(* Logix 5000 project; controller TFF vendor 1 type 14 code 107 rev 34.11; software revision 34.03; part 28 of 36 *)
(* tags used below, declared in another part *)
   Config : Configuration;   // Index Array used in configuration routines
   AlarmControl : AlarmControl;   // Alarm Control
   AnalogOutput : AnalogOutput[25];   // Analog Output Array
   AnalogPoint : AnalogInput[50];   // Analog Input Array
   CCPSystem : CCPSystem;   // CCP System Data
   ChartMark : ChartMark;   // Chart Mark
   Concentration : Concentration;
   CPU_Scanning : BOOL;   // System Scanning Flag
   Diafiltration : Diafiltration;
   DigitalOutput : BOOL[256];   // Digital Output Array these bits are sent to output cards.
   DigitalPoint : DigitalPoint[150];   // Digital Point Array
   DPAlarm : ALIAS FOR AlarmAnalog[40];   // Differential Pressure Alarm
   Drive : Drive[11];   // Drives Array
   ES001 : ALIAS FOR DigitalPoint[3];   // Emergency Stop
   Feed_Pump_P001_Type : INT;   // Feed Pump P001 Type Status
   FirstScanComplete : BOOL;   // First Scan Complete Flag
   FlowPath : FlowPath[64];   // Flow Path Array
   Membrane_Data : Membrane_Data;   // Membrane Data
   Mixer : Mixer;   // Mixer config. structure
   OperatingTime : OperatingTime;
   Operation : Operation[6,251];   // Operation Table
   Options : Options;   // Options List
   Phase0 : ALIAS FOR Phase[0];   // Phase 0
   Phase0_Totalizer_Feed : ALIAS FOR PhaseTotalizer[0];   // Phase 0 Total Feed
   Phase0_Totalizer_Filtrate : ALIAS FOR PhaseTotalizer[6];   // Phase 0 Total Filtrate
   Phase0_Totalizer_Retentate : ALIAS FOR PhaseTotalizer[12];   // Phase 0 Total Retentate
   PipeAnimation : PipeAnimation;   // HMI Pipe Animation Array
   PLCFault : FaultRecordType;   // PLC Major Fault Record
   PumpRunStatus : DINT;   // Pumps Run Status (1 = At least one pump running , 0 = no pump running)
   Rack_Murr_Node6_IND331_WI001 : IO_Station;   // Status of Node 6 IND331 WI001
   Rack_Murr_Node7_IND131_WI101 : IO_Station;   // Status of Node 7 IND131 WI101
   SIC001 : ALIAS FOR Drive[1];   // Feed Pump
   SIC002 : ALIAS FOR Drive[2];   // Transfer Pump
   SIC003 : ALIAS FOR Drive[3];   // Mixer
   SIC003DF : ALIAS FOR DigitalPoint[14];   // Mixer Defect
   SysControl : SysControl;   // General system status and command
   Tank : TankManagement;   // Tank Management
   ThisSystem : SystemType;
   TimerControl : TimerControl;   // Timer Control
   Timers : Timers[22];   // Timer Array
   TMPAlarm : ALIAS FOR AlarmAnalog[41];   // Trans-membrane Pressure Alarm
   Totalizer : Totalizers[20];   // Totalizers Array
   Transfer_Pump_P002_Type : INT;   // Transfer Pump P002 Type Status
   UserAlarm : UserAlarm;   // User Alarm (used in CCP Recipe)
   UserCr1 : ALIAS FOR DigitalPoint[65];   // User Critical Alarm 1
   UserCr2 : ALIAS FOR DigitalPoint[67];   // User Critical Alarm 2
   UserNCr1 : ALIAS FOR DigitalPoint[64];   // User Non Critical Alarm 1
   UserNCr2 : ALIAS FOR DigitalPoint[66];   // User Non Critical Alarm 2
   UserTime : ALIAS FOR Timers[18];   // User time
   UserTotalizerManagement : UserTotalizerManagement;   // User Totalizer management
   Valve : Valve[100];   // Valve Array
   XC102_3 : ALIAS FOR DigitalOutput[5];   // UV Auto Zero
   XS011 : ALIAS FOR DigitalPoint[11];   // Pump P001 Type
   XS012 : ALIAS FOR DigitalPoint[12];   // Pump P002 Type
   YA10 : ALIAS FOR DigitalPoint[59];   // PLC Program Major Fault
   YA41 : ALIAS FOR DigitalPoint[77];   // YA41 Operating Time Exceeded
(* Process, continued *)

ROUTINE InputProcessing   (* ladder *)
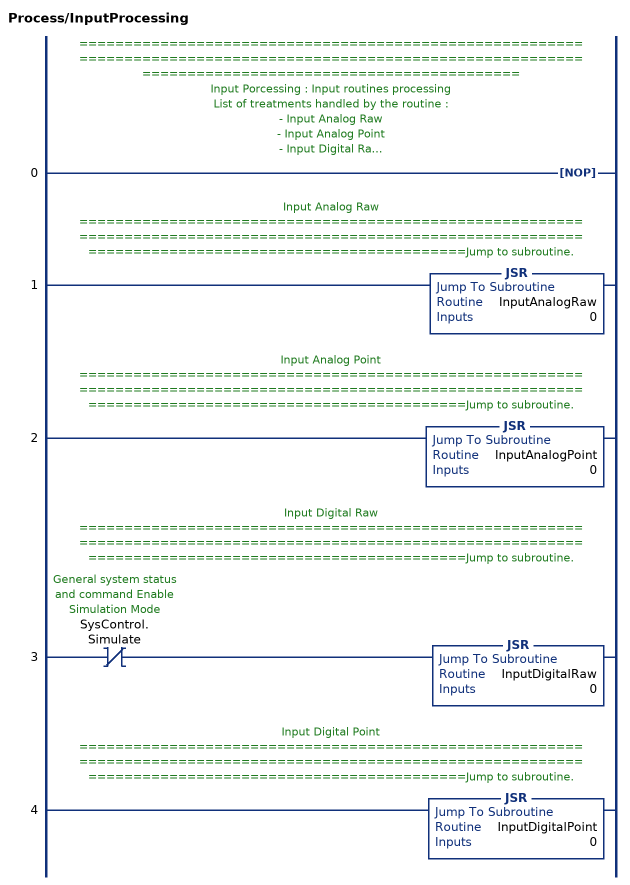
   // ==========================================================================================================================================================
   //                                                                                                                      Input Porcessing : Input routines processing
   //                                                     List of treatments handled by the routine :
   //                                                          - Input Analog Raw
   //                                                          - Input Analog Point
   //                                                          - Input Digital Raw
   //                                                          - Input Digital Point
   //                                                     -----------------------------------------------------------------------------------------------------------------------------------------------------
   //                                                     History
   //                                                          2019-AUG-13 - Actemium - B. Roch - Initial version for Candidate Release 3.00.00.00.a
   // ==========================================================================================================================================================
   0: NOP();
   // Input Analog Raw
   // ==========================================================================================================================================================Jump to subroutine.
   1: JSR(InputAnalogRaw,0);
   // Input Analog Point
   // ==========================================================================================================================================================Jump to subroutine.
   2: JSR(InputAnalogPoint,0);
   // Input Digital Raw
   // ==========================================================================================================================================================Jump to subroutine.
   3: XIO(SysControl.Simulate)JSR(InputDigitalRaw,0);
   // Input Digital Point
   // ==========================================================================================================================================================Jump to subroutine.
   4: JSR(InputDigitalPoint,0);
END_ROUTINE

ROUTINE MainRoutine   (* ladder *)
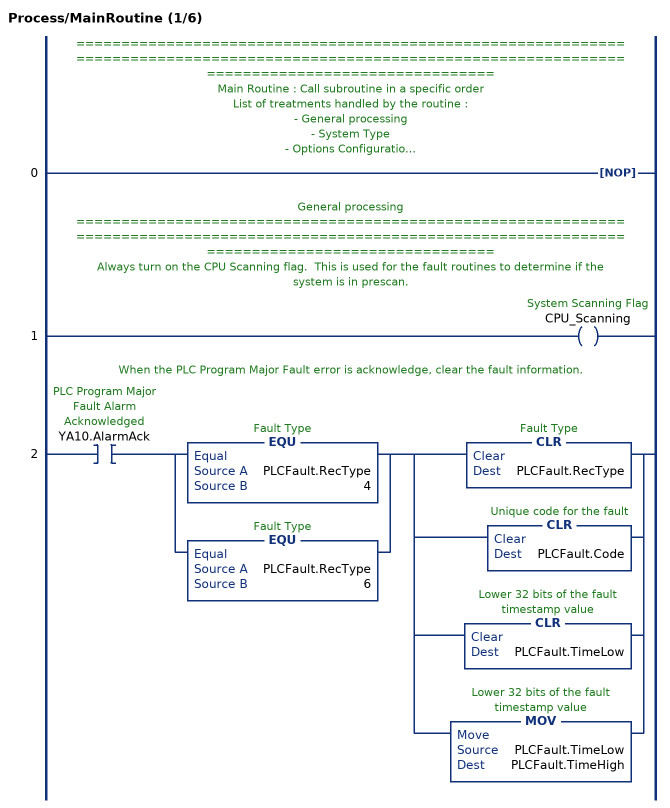
   // ==========================================================================================================================================================
   //                                                                                                            Main Routine : Call subroutine in a specific order
   //                                                     List of treatments handled by the routine :
   //                                                          - General processing
   //                                                          - System Type
   //                                                          - Options Configuration
   //                                                          - AnalogOutput Configuration
   //                                                          - AnalogPoint Configuration
   //                                                          - DigitalPoint Configuration (real input)
   //                                                          - DigitalPoint Configuration (soft input)
   //                                                          - Valve Configuration
   //                                                          - Drive Configuration
   //                                                          - Control Loop Configuration
   //                                                          - Totalizers Configuration
   //                                                          - Flowpath Configuration
   //                                                          - Reset Configuration
   //                                                          - Station Status
   //                                                          - Derived Data
   //                                                          - Analog and Digital Input Processing
   //                                                          - Pump Control
   //                                                          - Loop Control
   //                                                          - Valve Control
   //                                                          - Pipe Animation
   //                                                          - Alarm
   //                                                          - Concentration & Diafiltration
   //                                                          - TankManagement
   //                                                          - Miscellaneous Functions
   //                                                          - Analog and Digital Output Processing
   //                                                     -----------------------------------------------------------------------------------------------------------------------------------------------------
   //                                                     History
   //                                                          2019-AUG-13 - Actemium - B. Roch - Initial version for Candidate Release 3.00.00.00.a
   //                                                          2020-SEP-14 - Merck - Q. Spindler - Modifications for Candidate Release 3.00.00.01.a
   //                                                                  - Add TimerControl.TickMainTask for 1 sec tick in Main task
   // ==========================================================================================================================================================
   0: NOP();
   // General processing
   // ==========================================================================================================================================================
   // Always turn on the CPU Scanning flag.  This is used for the fault routines to determine if the system is in prescan.
   1: OTE(CPU_Scanning);
   // When the PLC Program Major Fault error is acknowledge, clear the fault information.
   2: XIC(YA10.AlarmAck)[EQU(PLCFault.RecType,4) ,EQU(PLCFault.RecType,6) ][CLR(PLCFault.RecType) ,CLR(PLCFault.Code) ,CLR(PLCFault.TimeLow) ,MOV(PLCFault.TimeLow,PLCFault.TimeHigh) ];
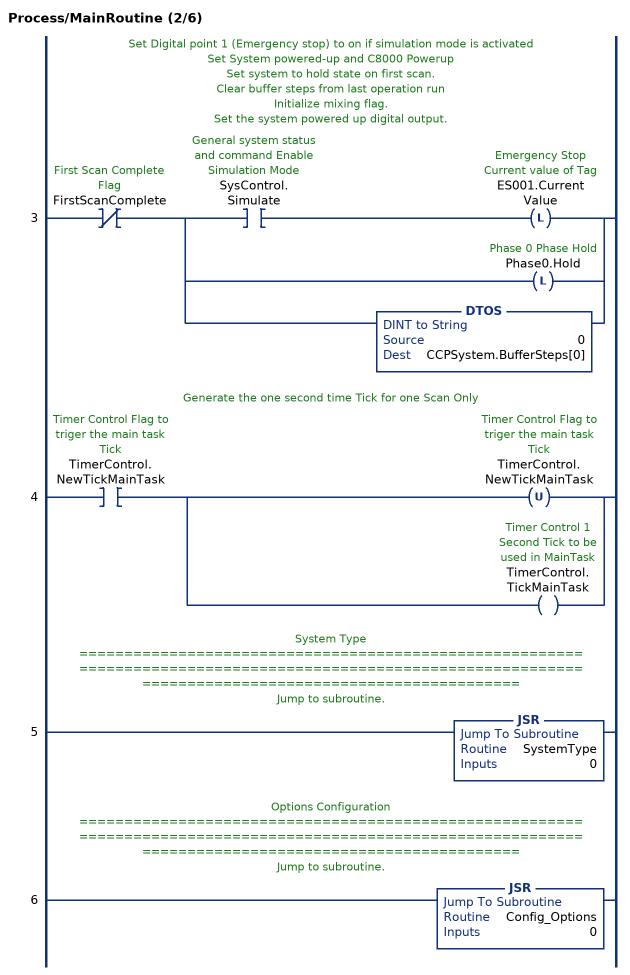
   // Set Digital point 1 (Emergency stop) to on if simulation mode is activated
   // Set System powered-up and C8000 Powerup
   // Set system to hold state on first scan.
   // Clear buffer steps from last operation run
   // Initialize mixing flag.
   // Set the system powered up digital output.
   3: XIO(FirstScanComplete)[XIC(SysControl.Simulate) OTL(ES001.CurrentValue) ,OTL(Phase0.Hold) ,DTOS(0,CCPSystem.BufferSteps[0]) ];
   // Generate the one second time Tick for one Scan Only
   4: XIC(TimerControl.NewTickMainTask)[OTU(TimerControl.NewTickMainTask) ,OTE(TimerControl.TickMainTask) ];
   // System Type
   // ==========================================================================================================================================================
   // Jump to subroutine.
   5: JSR(SystemType,0);
   // Options Configuration
   // ==========================================================================================================================================================
   // Jump to subroutine.
   6: JSR(Config_Options,0);
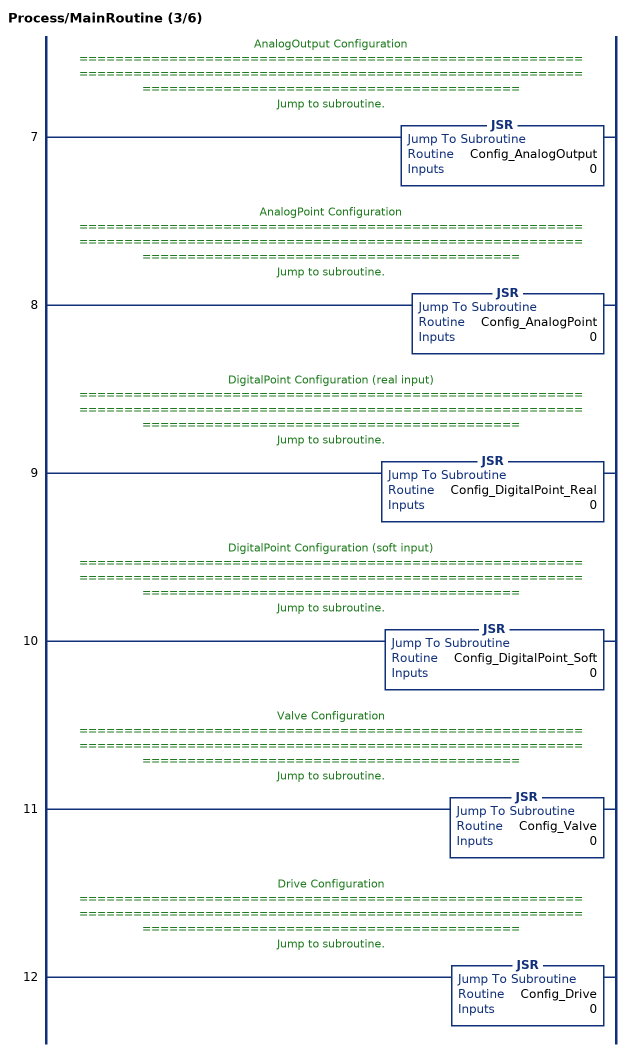
   // AnalogOutput Configuration
   // ==========================================================================================================================================================
   // Jump to subroutine.
   7: JSR(Config_AnalogOutput,0);
   // AnalogPoint Configuration
   // ==========================================================================================================================================================
   // Jump to subroutine.
   8: JSR(Config_AnalogPoint,0);
   // DigitalPoint Configuration (real input)
   // ==========================================================================================================================================================
   // Jump to subroutine.
   9: JSR(Config_DigitalPoint_Real,0);
   // DigitalPoint Configuration (soft input)
   // ==========================================================================================================================================================
   // Jump to subroutine.
   10: JSR(Config_DigitalPoint_Soft,0);
   // Valve Configuration
   // ==========================================================================================================================================================
   // Jump to subroutine.
   11: JSR(Config_Valve,0);
   // Drive Configuration
   // ==========================================================================================================================================================
   // Jump to subroutine.
   12: JSR(Config_Drive,0);
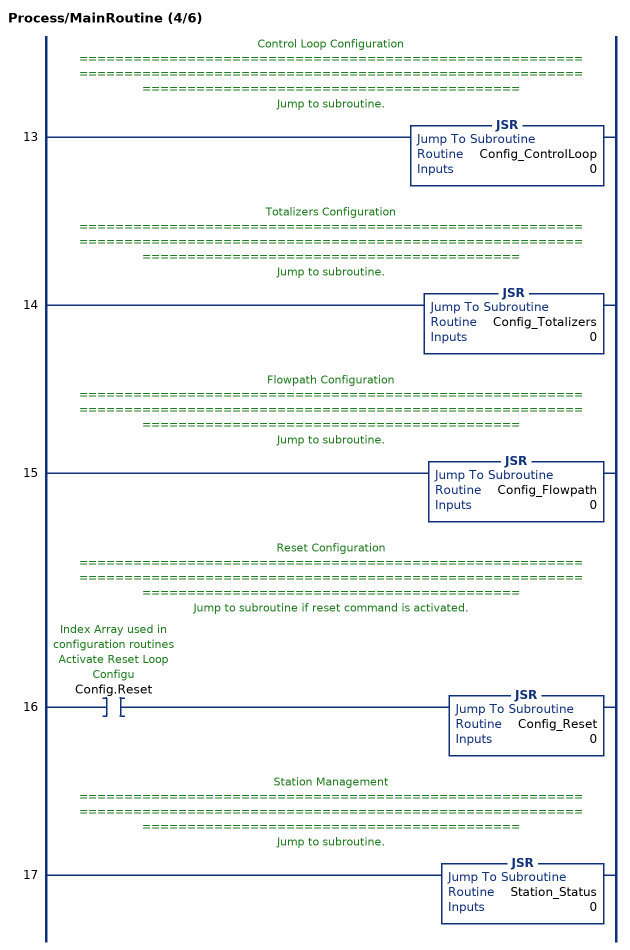
   // Control Loop Configuration
   // ==========================================================================================================================================================
   // Jump to subroutine.
   13: JSR(Config_ControlLoop,0);
   // Totalizers Configuration
   // ==========================================================================================================================================================
   // Jump to subroutine.
   14: JSR(Config_Totalizers,0);
   // Flowpath Configuration
   // ==========================================================================================================================================================
   // Jump to subroutine.
   15: JSR(Config_Flowpath,0);
   // Reset Configuration
   // ==========================================================================================================================================================
   // Jump to subroutine if reset command is activated.
   16: XIC(Config.Reset)JSR(Config_Reset,0);
   // Station Management
   // ==========================================================================================================================================================
   // Jump to subroutine.
   17: JSR(Station_Status,0);
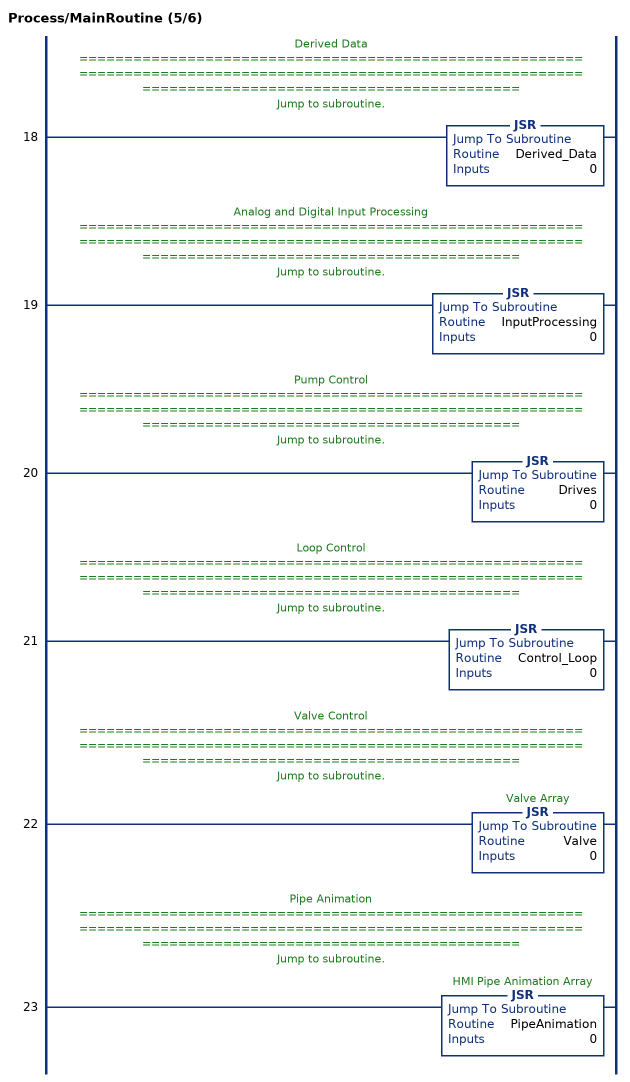
   // Derived Data
   // ==========================================================================================================================================================
   // Jump to subroutine.
   18: JSR(Derived_Data,0);
   // Analog and Digital Input Processing
   // ==========================================================================================================================================================
   // Jump to subroutine.
   19: JSR(InputProcessing,0);
   // Pump Control
   // ==========================================================================================================================================================
   // Jump to subroutine.
   20: JSR(Drives,0);
   // Loop Control
   // ==========================================================================================================================================================
   // Jump to subroutine.
   21: JSR(Control_Loop,0);
   // Valve Control
   // ==========================================================================================================================================================
   // Jump to subroutine.
   22: JSR(Valve,0);
   // Pipe Animation
   // ==========================================================================================================================================================
   // Jump to subroutine.
   23: JSR(PipeAnimation,0);
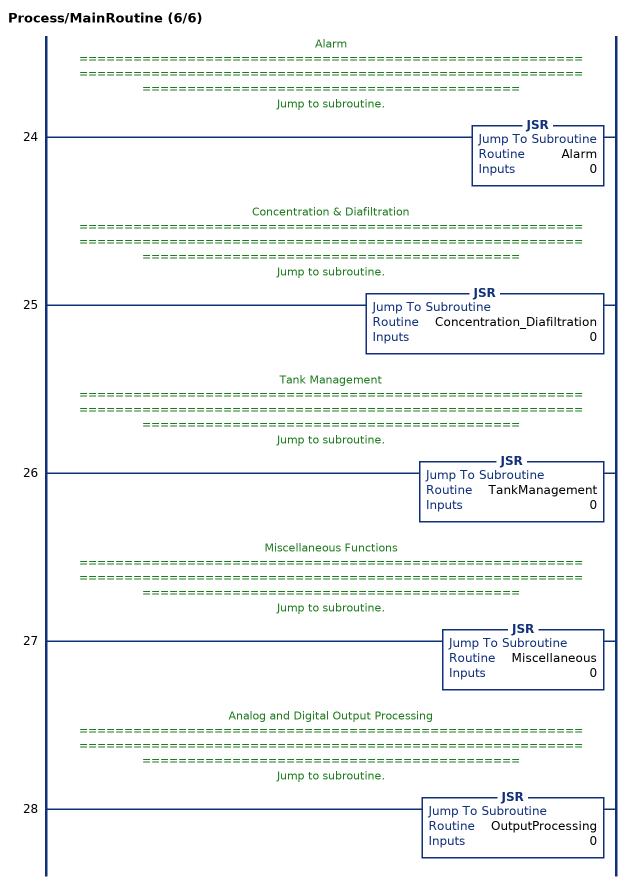
   // Alarm
   // ==========================================================================================================================================================
   // Jump to subroutine.
   24: JSR(Alarm,0);
   // Concentration & Diafiltration
   // ==========================================================================================================================================================
   // Jump to subroutine.
   25: JSR(Concentration_Diafiltration,0);
   // Tank Management
   // ==========================================================================================================================================================
   // Jump to subroutine.
   26: JSR(TankManagement,0);
   // Miscellaneous Functions
   // ==========================================================================================================================================================
   // Jump to subroutine.
   27: JSR(Miscellaneous,0);
   // Analog and Digital Output Processing
   // ==========================================================================================================================================================
   // Jump to subroutine.
   28: JSR(OutputProcessing,0);
END_ROUTINE

ROUTINE Miscellaneous   (* ladder *)
// Miscellaneous Routine
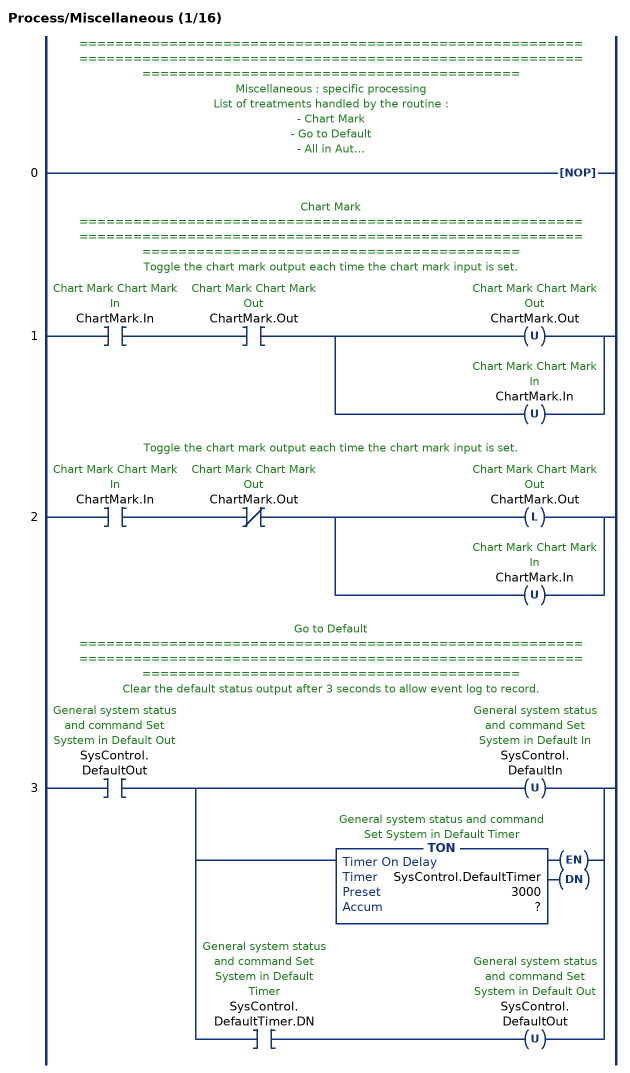
   // ==========================================================================================================================================================
   //                                                                                                                                 Miscellaneous : specific processing
   //                                                     List of treatments handled by the routine :
   //                                                          - Chart Mark
   //                                                          - Go to Default
   //                                                          - All in Auto
   //                                                          - Input Digital Point
   //                                                          - Enable All Alarms
   //                                                          - Disable All Alarms
   //                                                          - Enable all Analog signal alarms
   //                                                          - Disable all Analog signal alarms
   //                                                          - User totalizer management
   //                                                          - Pump Status calculation
   //                                                          - User Alarm (used in recipe only)
   //                                                          - Default Status
   //                                                          - Save \ Restore parameters conditions
   //                                                          - Mixer Reset Alarm Command
   //                                                          - IND331 and IND131 Configurations
   //                                                          - UV Baseline Zero Command Logic
   //                                                          - Pump Type Status
   //                                                     -----------------------------------------------------------------------------------------------------------------------------------------------------
   //                                                     History
   //                                                          2019-AUG-13 - Actemium - B. Roch - Initial version for Candidate Release 3.00.00.00.a
   //                                                          2019-OCT-25 - Actemium - B. Roch - Modification for Candidate Release 3.00.00.00.d
   //                                                         - Change Mixer Reset alarm condition SIC003DF.CurrentValue instead of SIC003DF.Alarm
   //                                                      2020-SEP-29 - Merck - Q. Spindler - Modifications for Candidate Release 3.00.00.01.a
   // 							- Add Retentate totalizer for UserTotalizer
   //                                                             2021-APR-30 - DAVIDSON- Ch. ARBOGAST - Modifications for Candidate Release 3.01.00.00.a
   //             -  Add Conditions to YA41 Operating Time Exceeded
   // ==========================================================================================================================================================
   0: NOP();
   // Chart Mark
   // ==========================================================================================================================================================
   // Toggle the chart mark output each time the chart mark input is set.
   1: XIC(ChartMark.In)XIC(ChartMark.Out)[OTU(ChartMark.Out) ,OTU(ChartMark.In) ];
   // Toggle the chart mark output each time the chart mark input is set.
   2: XIC(ChartMark.In)XIO(ChartMark.Out)[OTL(ChartMark.Out) ,OTU(ChartMark.In) ];
   // Go to Default
   // ==========================================================================================================================================================
   // Clear the default status output after 3 seconds to allow event log to record.
   3: XIC(SysControl.DefaultOut)[OTU(SysControl.DefaultIn) ,TON(SysControl.DefaultTimer,?,?) ,XIC(SysControl.DefaultTimer.DN) OTU(SysControl.DefaultOut) ];
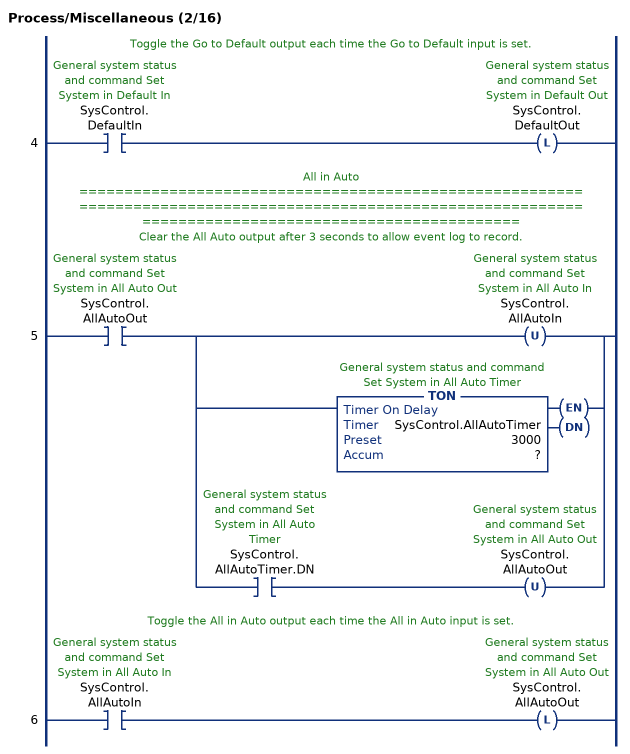
   // Toggle the Go to Default output each time the Go to Default input is set.
   4: XIC(SysControl.DefaultIn)OTL(SysControl.DefaultOut);
   // All in Auto
   // ==========================================================================================================================================================
   // Clear the All Auto output after 3 seconds to allow event log to record.
   5: XIC(SysControl.AllAutoOut)[OTU(SysControl.AllAutoIn) ,TON(SysControl.AllAutoTimer,?,?) ,XIC(SysControl.AllAutoTimer.DN) OTU(SysControl.AllAutoOut) ];
   // Toggle the All in Auto output each time the All in Auto input is set.
   6: XIC(SysControl.AllAutoIn)OTL(SysControl.AllAutoOut);
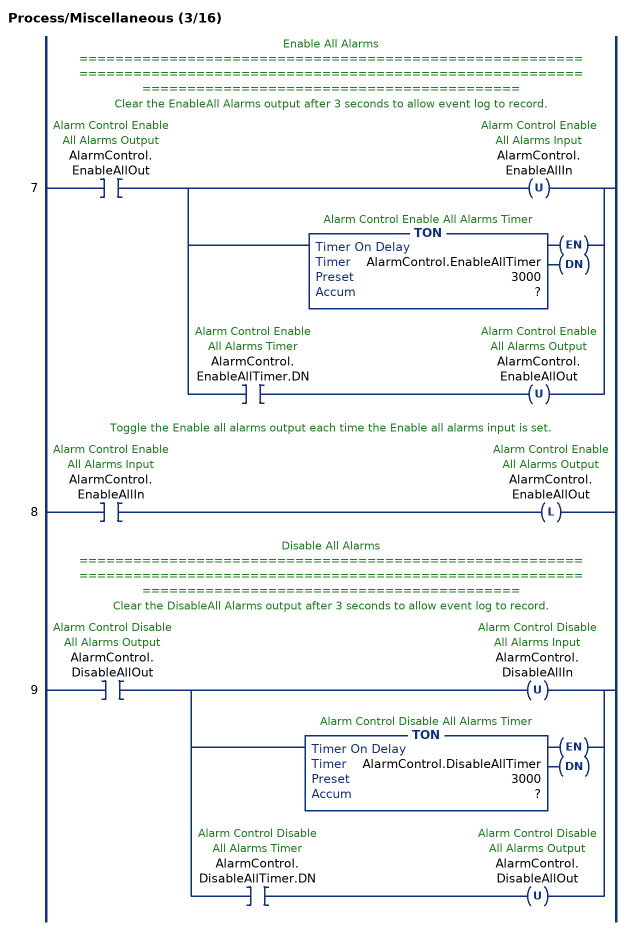
   // Enable All Alarms
   // ==========================================================================================================================================================
   // Clear the EnableAll Alarms output after 3 seconds to allow event log to record.
   7: XIC(AlarmControl.EnableAllOut)[OTU(AlarmControl.EnableAllIn) ,TON(AlarmControl.EnableAllTimer,?,?) ,XIC(AlarmControl.EnableAllTimer.DN) OTU(AlarmControl.EnableAllOut) ];
   // Toggle the Enable all alarms output each time the Enable all alarms input is set.
   8: XIC(AlarmControl.EnableAllIn)OTL(AlarmControl.EnableAllOut);
   // Disable All Alarms
   // ==========================================================================================================================================================
   // Clear the DisableAll Alarms output after 3 seconds to allow event log to record.
   9: XIC(AlarmControl.DisableAllOut)[OTU(AlarmControl.DisableAllIn) ,TON(AlarmControl.DisableAllTimer,?,?) ,XIC(AlarmControl.DisableAllTimer.DN) OTU(AlarmControl.DisableAllOut) ];
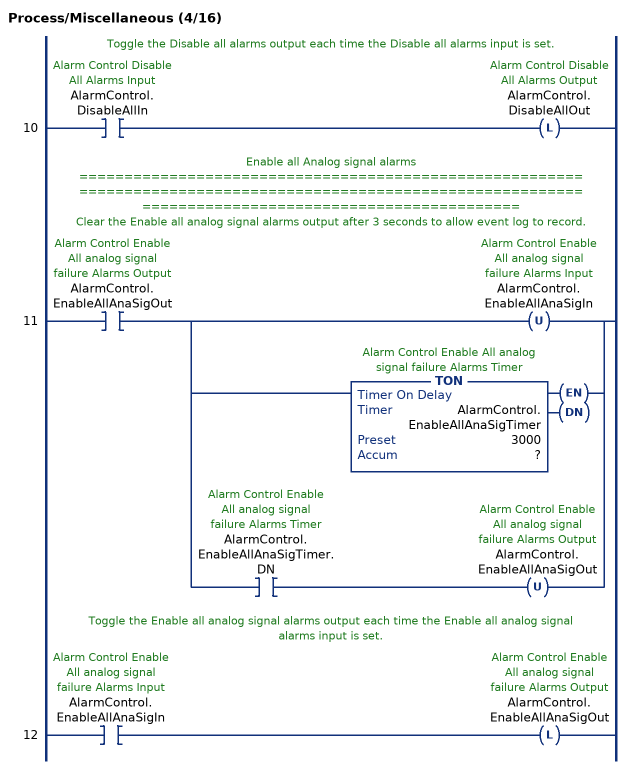
   // Toggle the Disable all alarms output each time the Disable all alarms input is set.
   10: XIC(AlarmControl.DisableAllIn)OTL(AlarmControl.DisableAllOut);
   // Enable all Analog signal alarms
   // ==========================================================================================================================================================
   // Clear the Enable all analog signal alarms output after 3 seconds to allow event log to record.
   11: XIC(AlarmControl.EnableAllAnaSigOut)[OTU(AlarmControl.EnableAllAnaSigIn) ,TON(AlarmControl.EnableAllAnaSigTimer,?,?) ,XIC(AlarmControl.EnableAllAnaSigTimer.DN) OTU(AlarmControl.EnableAllAnaSigOut) ];
   // Toggle the Enable all analog signal alarms output each time the Enable all analog signal alarms input is set.
   12: XIC(AlarmControl.EnableAllAnaSigIn)OTL(AlarmControl.EnableAllAnaSigOut);
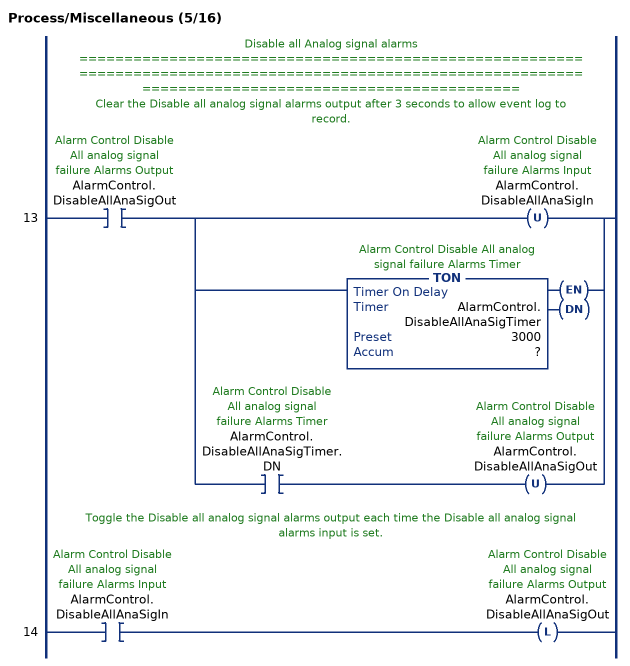
   // Disable all Analog signal alarms
   // ==========================================================================================================================================================
   // Clear the Disable all analog signal alarms output after 3 seconds to allow event log to record.
   13: XIC(AlarmControl.DisableAllAnaSigOut)[OTU(AlarmControl.DisableAllAnaSigIn) ,TON(AlarmControl.DisableAllAnaSigTimer,?,?) ,XIC(AlarmControl.DisableAllAnaSigTimer.DN) OTU(AlarmControl.DisableAllAnaSigOut) ];
   // Toggle the Disable all analog signal alarms output each time the Disable all analog signal alarms input is set.
   14: XIC(AlarmControl.DisableAllAnaSigIn)OTL(AlarmControl.DisableAllAnaSigOut);
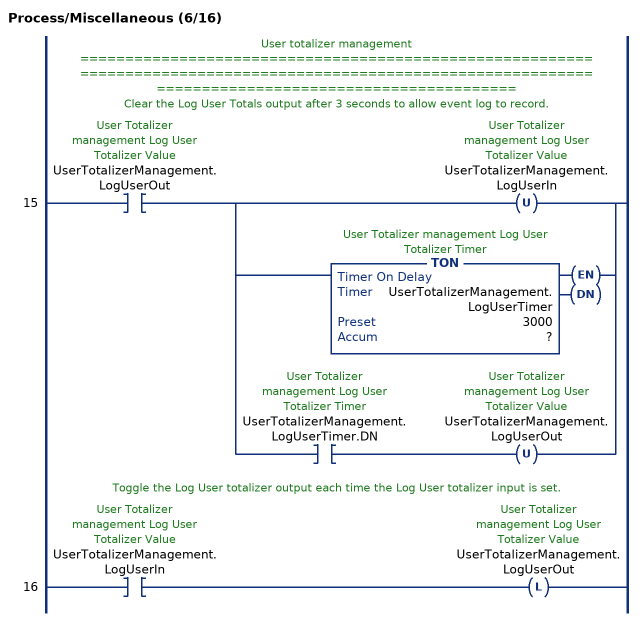
   // User totalizer management
   // ==========================================================================================================================================================
   // Clear the Log User Totals output after 3 seconds to allow event log to record.
   15: XIC(UserTotalizerManagement.LogUserOut)[OTU(UserTotalizerManagement.LogUserIn) ,TON(UserTotalizerManagement.LogUserTimer,?,?) ,XIC(UserTotalizerManagement.LogUserTimer.DN) OTU(UserTotalizerManagement.LogUserOut) ];
   // Toggle the Log User totalizer output each time the Log User totalizer input is set.
   16: XIC(UserTotalizerManagement.LogUserIn)OTL(UserTotalizerManagement.LogUserOut);
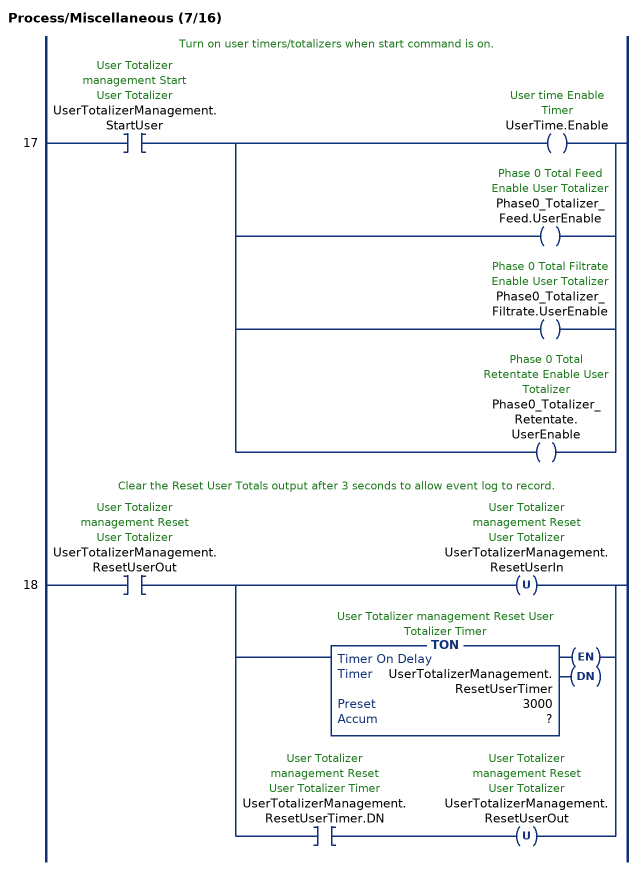
   // Turn on user timers/totalizers when start command is on.
   17: XIC(UserTotalizerManagement.StartUser)[OTE(UserTime.Enable) ,OTE(Phase0_Totalizer_Feed.UserEnable) ,OTE(Phase0_Totalizer_Filtrate.UserEnable) ,OTE(Phase0_Totalizer_Retentate.UserEnable) ];
   // Clear the Reset User Totals output after 3 seconds to allow event log to record.
   18: XIC(UserTotalizerManagement.ResetUserOut)[OTU(UserTotalizerManagement.ResetUserIn) ,TON(UserTotalizerManagement.ResetUserTimer,?,?) ,XIC(UserTotalizerManagement.ResetUserTimer.DN) OTU(UserTotalizerManagement.ResetUserOut) ];
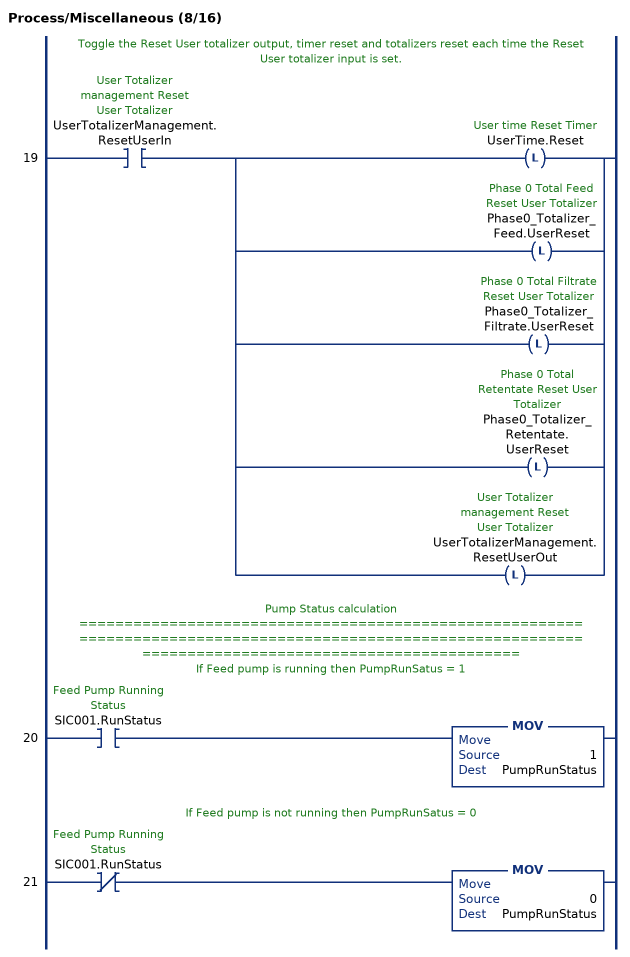
   // Toggle the Reset User totalizer output, timer reset and totalizers reset each time the Reset User totalizer input is set.
   19: XIC(UserTotalizerManagement.ResetUserIn)[OTL(UserTime.Reset) ,OTL(Phase0_Totalizer_Feed.UserReset) ,OTL(Phase0_Totalizer_Filtrate.UserReset) ,OTL(Phase0_Totalizer_Retentate.UserReset) ,OTL(UserTotalizerManagement.ResetUserOut) ];
   // Pump Status calculation
   // ==========================================================================================================================================================
   // If Feed pump is running then PumpRunSatus = 1
   20: XIC(SIC001.RunStatus)MOV(1,PumpRunStatus);
   // If Feed pump is not running then PumpRunSatus = 0
   21: XIO(SIC001.RunStatus)MOV(0,PumpRunStatus);
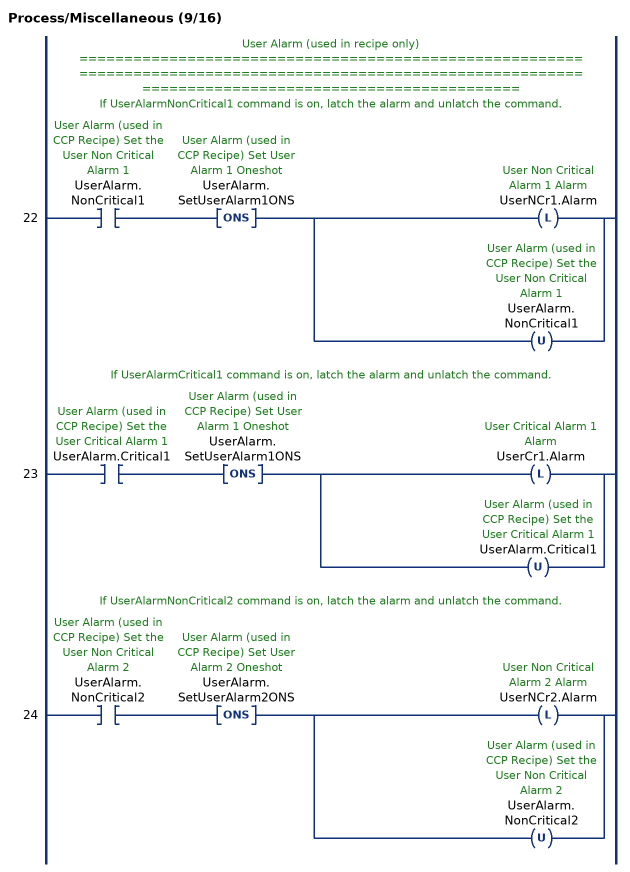
   // User Alarm (used in recipe only)
   // ==========================================================================================================================================================
   // If UserAlarmNonCritical1 command is on, latch the alarm and unlatch the command.
   22: XIC(UserAlarm.NonCritical1)ONS(UserAlarm.SetUserAlarm1ONS)[OTL(UserNCr1.Alarm) ,OTU(UserAlarm.NonCritical1) ];
   // If UserAlarmCritical1 command is on, latch the alarm and unlatch the command.
   23: XIC(UserAlarm.Critical1)ONS(UserAlarm.SetUserAlarm1ONS)[OTL(UserCr1.Alarm) ,OTU(UserAlarm.Critical1) ];
   // If UserAlarmNonCritical2 command is on, latch the alarm and unlatch the command.
   24: XIC(UserAlarm.NonCritical2)ONS(UserAlarm.SetUserAlarm2ONS)[OTL(UserNCr2.Alarm) ,OTU(UserAlarm.NonCritical2) ];
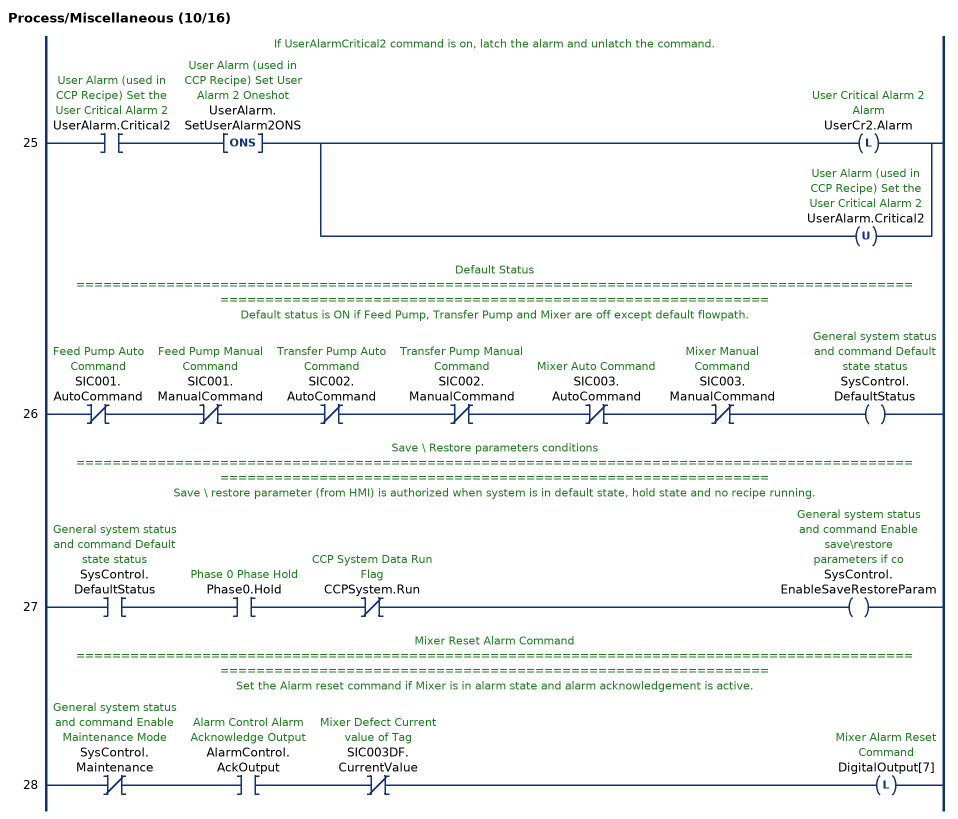
   // If UserAlarmCritical2 command is on, latch the alarm and unlatch the command.
   25: XIC(UserAlarm.Critical2)ONS(UserAlarm.SetUserAlarm2ONS)[OTL(UserCr2.Alarm) ,OTU(UserAlarm.Critical2) ];
   // Default Status
   // ==========================================================================================================================================================
   // Default status is ON if Feed Pump, Transfer Pump and Mixer are off except default flowpath.
   26: XIO(SIC001.AutoCommand)XIO(SIC001.ManualCommand)XIO(SIC002.AutoCommand)XIO(SIC002.ManualCommand)XIO(SIC003.AutoCommand)XIO(SIC003.ManualCommand)OTE(SysControl.DefaultStatus);
   // Save \ Restore parameters conditions
   // ==========================================================================================================================================================
   // Save \ restore parameter (from HMI) is authorized when system is in default state, hold state and no recipe running.
   27: XIC(SysControl.DefaultStatus)XIC(Phase0.Hold)XIO(CCPSystem.Run)OTE(SysControl.EnableSaveRestoreParam);
   // Mixer Reset Alarm Command
   // ==========================================================================================================================================================
   // Set the Alarm reset command if Mixer is in alarm state and alarm acknowledgement is active.
   28: XIO(SysControl.Maintenance)XIC(AlarmControl.AckOutput)XIO(SIC003DF.CurrentValue)OTL(DigitalOutput[7]);
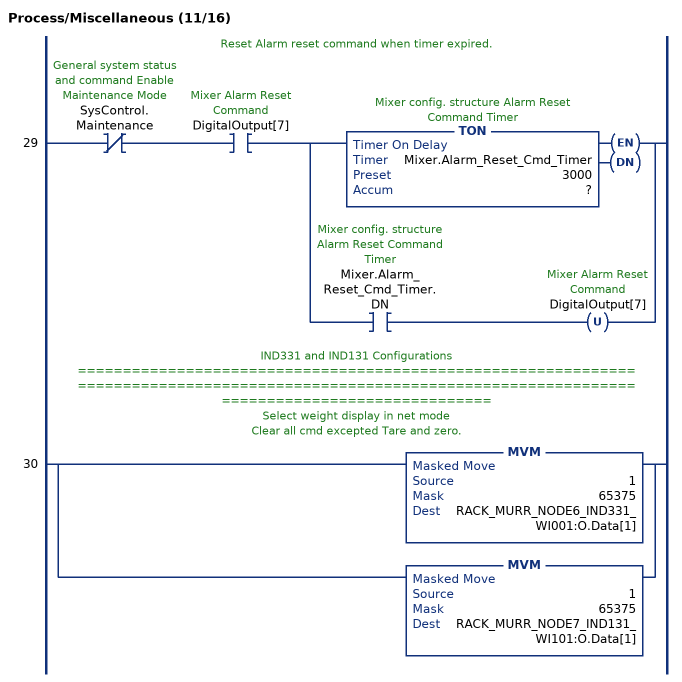
   // Reset Alarm reset command when timer expired.
   29: XIO(SysControl.Maintenance)XIC(DigitalOutput[7])[TON(Mixer.Alarm_Reset_Cmd_Timer,?,?) ,XIC(Mixer.Alarm_Reset_Cmd_Timer.DN) OTU(DigitalOutput[7]) ];
   // IND331 and IND131 Configurations
   // ==========================================================================================================================================================
   // Select weight display in net mode
   // Clear all cmd excepted Tare and zero.
   30: [MVM(1,65375,RACK_MURR_NODE6_IND331_WI001:O.Data[1]) ,MVM(1,65375,RACK_MURR_NODE7_IND131_WI101:O.Data[1]) ];
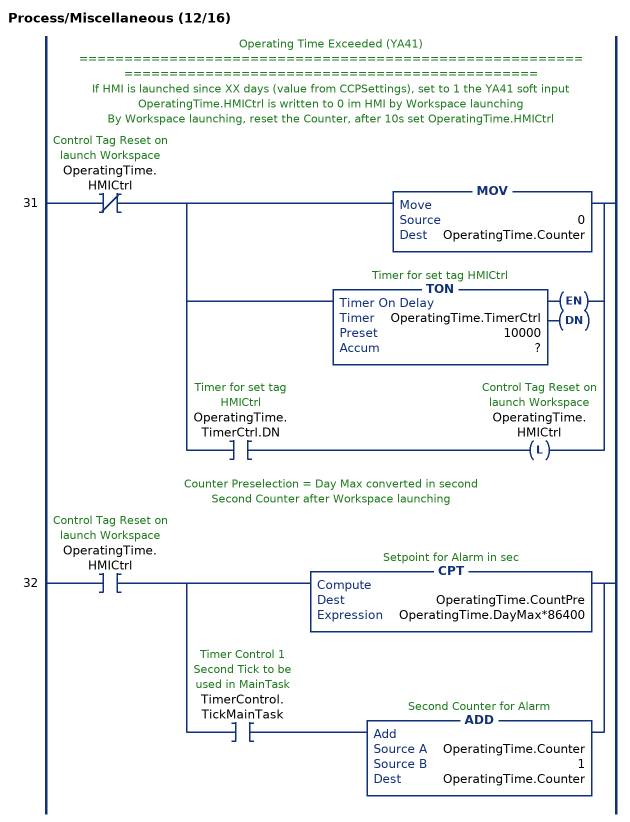
   // Operating Time Exceeded (YA41)
   // ======================================================================================================
   // If HMI is launched since XX days (value from CCPSettings), set to 1 the YA41 soft input
   // OperatingTime.HMICtrl is written to 0 im HMI by Workspace launching
   // By Workspace launching, reset the Counter, after 10s set OperatingTime.HMICtrl
   31: XIO(OperatingTime.HMICtrl)[MOV(0,OperatingTime.Counter) ,TON(OperatingTime.TimerCtrl,?,?) ,XIC(OperatingTime.TimerCtrl.DN) OTL(OperatingTime.HMICtrl) ];
   // Counter Preselection = Day Max converted in second
   // Second Counter after Workspace launching
   32: XIC(OperatingTime.HMICtrl)[CPT(OperatingTime.CountPre,OperatingTime.DayMax*86400) ,XIC(TimerControl.TickMainTask) ADD(OperatingTime.Counter,1,OperatingTime.Counter) ];
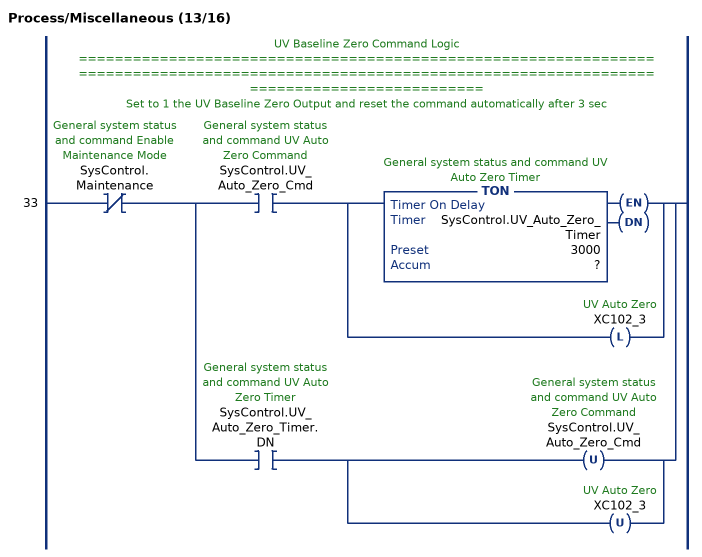
   // UV Baseline Zero Command Logic
   // ==========================================================================================================================================================
   // Set to 1 the UV Baseline Zero Output and reset the command automatically after 3 sec
   33: XIO(SysControl.Maintenance)[XIC(SysControl.UV_Auto_Zero_Cmd) [TON(SysControl.UV_Auto_Zero_Timer,?,?) ,OTL(XC102_3) ] ,XIC(SysControl.UV_Auto_Zero_Timer.DN) [OTU(SysControl.UV_Auto_Zero_Cmd) ,OTU(XC102_3) ] ];
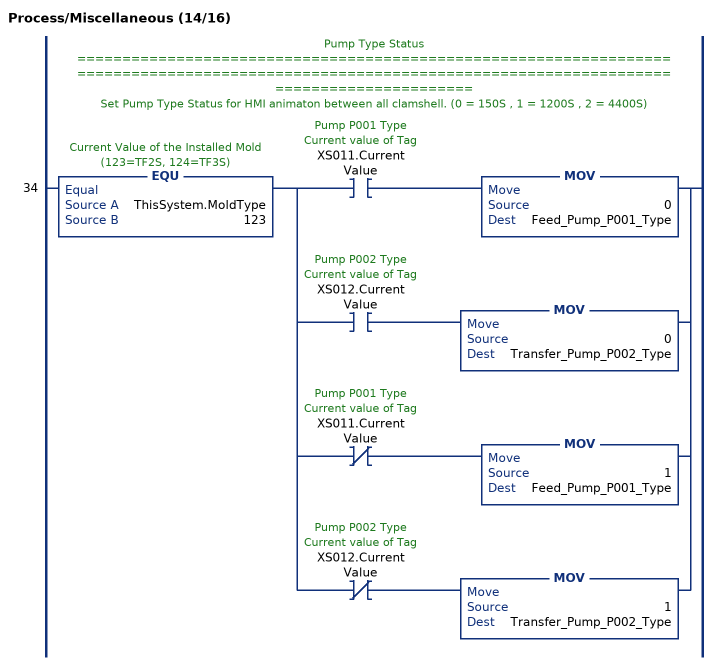
   // Pump Type Status
   // ==========================================================================================================================================================
   // Set Pump Type Status for HMI animaton between all clamshell. (0 = 150S , 1 = 1200S , 2 = 4400S)
   34: EQU(ThisSystem.MoldType,123)[XIC(XS011.CurrentValue) MOV(0,Feed_Pump_P001_Type) ,XIC(XS012.CurrentValue) MOV(0,Transfer_Pump_P002_Type) ,XIO(XS011.CurrentValue) MOV(1,Feed_Pump_P001_Type) ,XIO(XS012.CurrentValue) MOV(1,Transfer_Pump_P002_Type) ];
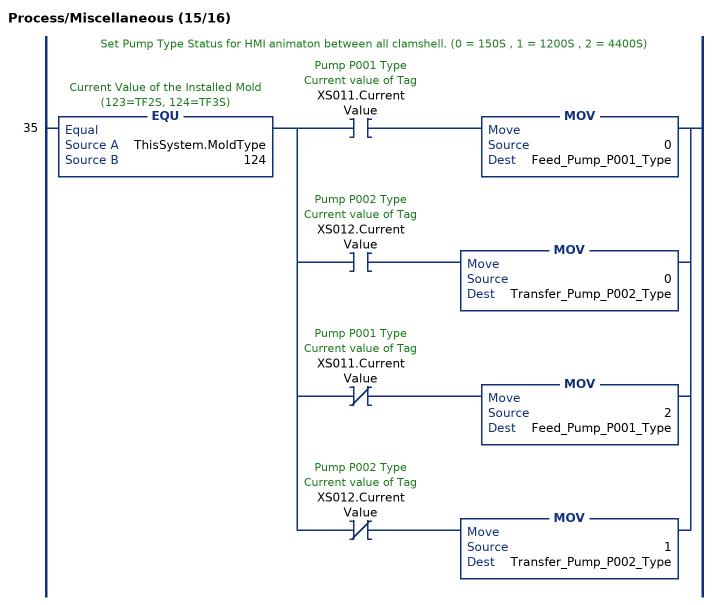
   // Set Pump Type Status for HMI animaton between all clamshell. (0 = 150S , 1 = 1200S , 2 = 4400S)
   35: EQU(ThisSystem.MoldType,124)[XIC(XS011.CurrentValue) MOV(0,Feed_Pump_P001_Type) ,XIC(XS012.CurrentValue) MOV(0,Transfer_Pump_P002_Type) ,XIO(XS011.CurrentValue) MOV(2,Feed_Pump_P001_Type) ,XIO(XS012.CurrentValue) MOV(1,Transfer_Pump_P002_Type) ];
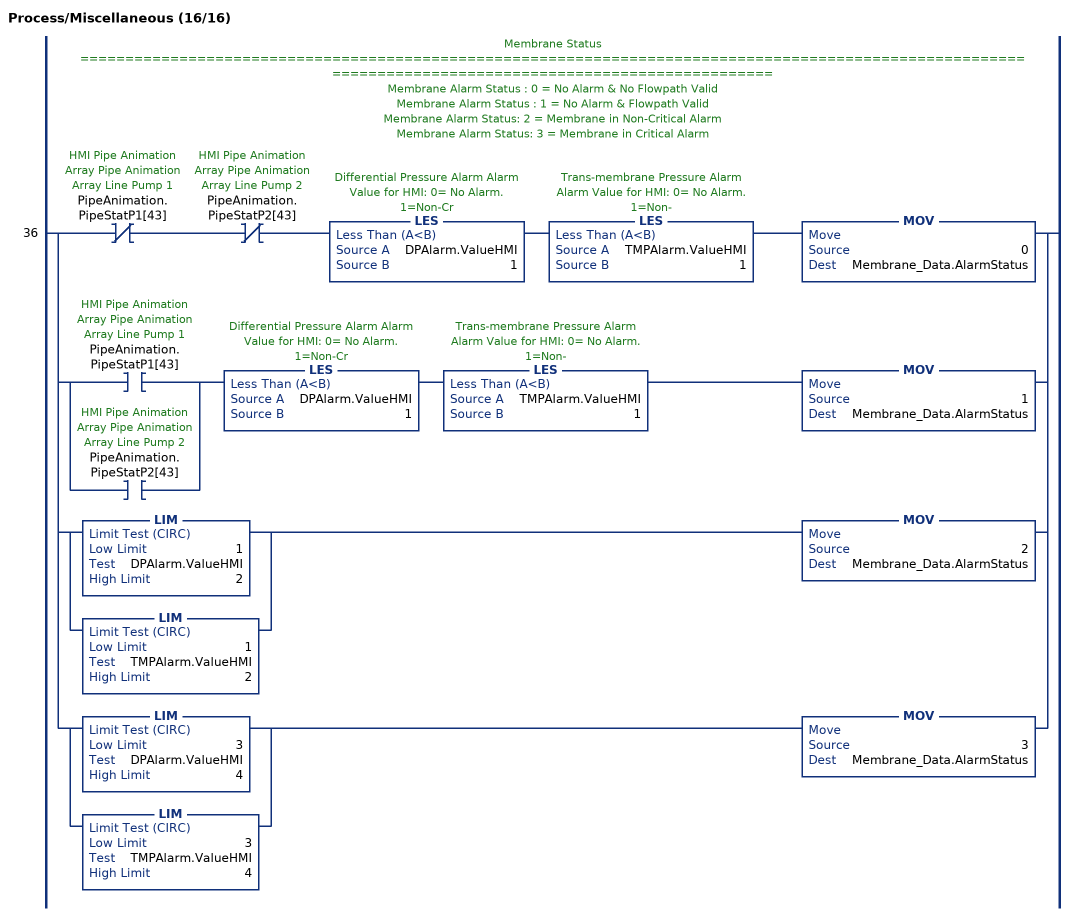
   // Membrane Status
   // ==========================================================================================================================================================
   // Membrane Alarm Status : 0 = No Alarm & No Flowpath Valid
   // Membrane Alarm Status : 1 = No Alarm & Flowpath Valid
   // Membrane Alarm Status: 2 = Membrane in Non-Critical Alarm
   // Membrane Alarm Status: 3 = Membrane in Critical Alarm
   36: [XIO(PipeAnimation.PipeStatP1[43]) XIO(PipeAnimation.PipeStatP2[43]) LES(DPAlarm.ValueHMI,1) LES(TMPAlarm.ValueHMI,1) MOV(0,Membrane_Data.AlarmStatus) ,[XIC(PipeAnimation.PipeStatP1[43]) ,XIC(PipeAnimation.PipeStatP2[43]) ] LES(DPAlarm.ValueHMI,1) LES(TMPAlarm.ValueHMI,1) MOV(1,Membrane_Data.AlarmStatus) ,[LIM(1,DPAlarm.ValueHMI,2) ,LIM(1,TMPAlarm.ValueHMI,2) ] MOV(2,Membrane_Data.AlarmStatus) ,[LIM(3,DPAlarm.ValueHMI,4) ,LIM(3,TMPAlarm.ValueHMI,4) ] MOV(3,Membrane_Data.AlarmStatus) ];
END_ROUTINE
